{attribute 'qualified_only'}
{attribute 'strict'}
TYPE E_CIP_ClientTank :
(
	eNone := 0,
	eClose,
	eTank_A,
	eTank_A_Sprinkler,
	eTank_B,
	eTank_B_Sprinkler,
	eDrain
);
END_TYPE

(* stored: Version 1.1.0.1, ProductVersion 3.1.4024.12
   DUT E_CIP_ClientTank: Id {a8ac13e7-a560-437e-9bbb-89d4cad6d00b} *)
